(* IEC 61131-3 sources: JingjiangArm/moonboxpro_arm_8.4/Application/Application/任务列表/CommTask/COMM_DIAMONDS/和金刚UDP通讯/功能接口, 6 files *)

(* ---- KS_CheckAll_StZone_UnSynchronized.st ---- *)
(*@CES
Name=KS_CheckAll_StZone_UnSynchronized
Type=FunctionBlock
TypeGuid=6f9dac99-8de1-4efc-8465-68ac443b7d08
Guid=07bfdfe8-2771-43fc-9a3c-80039394908a
HasDeclaration=True
HasImplementation=True
*)
{DECLARATION}
FUNCTION KS_CheckAll_StZone_UnSynchronized : INT(*0表示都同步了/>0表示未同步的数量/<0表示错误*)
VAR_INPUT
	i_pstStDataZone: POINTER TO StDataZone;(*读写区域*)
END_VAR
VAR
	uiN: UINT;
	iResult: INT;
END_VAR

{IMPLEMENTATION}
iResult:= 0;
IF i_pstStDataZone<>0 THEN
	FOR uiN:=1 TO i_pstStDataZone^.uiNodeNum BY 1 DO
		IF i_pstStDataZone^.astStDataNode[uiN].bySynchronized<>SINT_TO_BYTE(-1) THEN
			iResult:= iResult+1;(*未同步的数量+1*)
		END_IF
	END_FOR
ELSE
	iResult:= -1;
END_IF
KS_CheckAll_StZone_UnSynchronized:= iResult;

(* ---- KS_GenTxData_.st ---- *)
(*@CES
Name=KS_GenTxData_
Type=FunctionBlock
TypeGuid=6f9dac99-8de1-4efc-8465-68ac443b7d08
Guid=4f0cddb0-57bc-4748-9ef3-99d0df4ac11d
HasDeclaration=True
HasImplementation=True
*)
{DECLARATION}
FUNCTION KS_GenTxData_ : INT(*0无错误/-1参数非法/-100未支持的功能字/-200写多个寄存器范围无效*)
VAR_INPUT
	i_dwTxBuf: DWORD;
	i_pstStDataNode: POINTER TO StDataNode;
	i_dwBaseAdr: DWORD;
	i_uiInvocation: UINT;
	i_byFunctionId: BYTE;(*功能id/目前仅处理03和16*)
	i_piTxPayloadLen: POINTER TO INT;(*用于接收返回的实际tx数据数量/单位字节*)
	i_xOnlyWrite: BOOL;(*只写区域-16384*)
END_VAR
VAR
	iResult: INT := 0;
	uiTmp: UINT;
	pstStADU_tmp: POINTER TO StADU;
	pbyByteCount_tmp: POINTER TO BYTE;
	paiRegisters_tmp: POINTER TO ARRAY [1..MAX_PDU_REGISTERS] OF INT;
END_VAR
VAR CONSTANT
	MAX_PDU_REGISTERS: INT := 123;(*0X1~0X7B(最大)*)
	MB_FUNC_READ_MULTI_REGS: BYTE := 3;(*读多个寄存器*)
	MB_FUNC_WRITE_MULTI_REGS: BYTE := 16;(*写多个寄存器*)
END_VAR
{IMPLEMENTATION}
iResult:= 0;
IF i_dwTxBuf<>0 AND
	i_pstStDataNode<>0 AND
	i_piTxPayloadLen<>0 THEN

	(*主要的输入参数合法*)
	pstStADU_tmp:= i_dwTxBuf;

	(*mbap*)
	pstStADU_tmp^.stStMBAP.uiInvocation:= bswap_16(i_uiInvocation);
	pstStADU_tmp^.stStMBAP.uiProtocol:= 0;
	pstStADU_tmp^.stStMBAP.uiLength:= 0;(*这个长度根据i_byFunctionId的类别最后再重新统计比较合适*)
	pstStADU_tmp^.stStMBAP.byUnit:= 1;(*按slaveID=1/2025.8.4.192327*)

	(*pdu*)
	pstStADU_tmp^.stStPDU_Header.byFunction:= i_byFunctionId;
	IF i_byFunctionId=MB_FUNC_READ_MULTI_REGS THEN(*读多个寄存器*)
		(*功能字/单字节/不需要字序处理*)
		pstStADU_tmp^.stStPDU_Header.byFunction:= i_byFunctionId;

		(*地址和寄存器数量/16bit/都需要做字序处理*)
		pstStADU_tmp^.stStPDU_Header.uiAddress:= bswap_16(i_pstStDataNode^.uiAddress);
		pstStADU_tmp^.stStPDU_Header.uiQuantity:= bswap_16(i_pstStDataNode^.uiQuantity);

		(*更新mbap中的uiLength/16bit/需要处理字序*)
		uiTmp:= SIZEOF(pstStADU_tmp^.stStMBAP.byUnit) + SIZEOF(pstStADU_tmp^.stStPDU_Header);
		pstStADU_tmp^.stStMBAP.uiLength:= bswap_16(uiTmp);

		(*实际数据量*)
		i_piTxPayloadLen^:= DWORD_TO_INT(SIZEOF(pstStADU_tmp^));

	ELSIF i_byFunctionId=MB_FUNC_WRITE_MULTI_REGS THEN(*写多个寄存器*)
		(*功能字/单字节/不需要字序处理*)
		pstStADU_tmp^.stStPDU_Header.byFunction:= i_byFunctionId;

		(*地址和寄存器数量/16bit/都需要做字序处理*)
		IF i_pstStDataNode^.uiQuantity>=1 AND i_pstStDataNode^.uiQuantity<=MAX_PDU_REGISTERS THEN
			(*增加1级判断/保证寄存器在合法范围*)

			pstStADU_tmp^.stStPDU_Header.uiAddress:= bswap_16(i_pstStDataNode^.uiAddress);
			pstStADU_tmp^.stStPDU_Header.uiQuantity:= bswap_16(i_pstStDataNode^.uiQuantity);

			(*填充字节数量/单字节不用做字序处理*)
			pbyByteCount_tmp:= i_dwTxBuf + SIZEOF(pstStADU_tmp^);
			pbyByteCount_tmp^:= UINT_TO_BYTE(i_pstStDataNode^.uiQuantity*2);

			(*将寄存器数据搬到要发送的区域/这里没有做大小端数据处理*)
			paiRegisters_tmp:= i_dwTxBuf + SIZEOF(pstStADU_tmp^) + SIZEOF(pbyByteCount_tmp^);
			IF i_xOnlyWrite THEN
				SysMemCpy(
					paiRegisters_tmp,
					i_dwBaseAdr+(i_pstStDataNode^.uiAddress-PARAM_ZONE_C2S)*2,
					i_pstStDataNode^.uiQuantity*2);
			ELSE
				SysMemCpy(
					paiRegisters_tmp,
					i_dwBaseAdr+(i_pstStDataNode^.uiAddress-PARAM_ZONE_ALTERNATE_OFST)*2,
					i_pstStDataNode^.uiQuantity*2);
			END_IF

			(*更新mbap中的uiLength/16bit/需要处理字序*)
			uiTmp:= SIZEOF(pstStADU_tmp^.stStMBAP.byUnit) + SIZEOF(pstStADU_tmp^.stStPDU_Header) + SIZEOF(pbyByteCount_tmp^) + i_pstStDataNode^.uiQuantity*2;
			pstStADU_tmp^.stStMBAP.uiLength:= bswap_16(uiTmp);

			(*实际数据量*)
			i_piTxPayloadLen^:= DWORD_TO_INT(SIZEOF(pstStADU_tmp^) + SIZEOF(pbyByteCount_tmp^) + i_pstStDataNode^.uiQuantity*2);
		ELSE
			iResult:= -200;
		END_IF
	ELSE
		iResult:= -100;(*未支持的功能字*)
	END_IF
ELSE
	iResult:= -1;
END_IF
KS_GenTxData_:= iResult;

(* ---- KS_InitStProofList.st ---- *)
(*@CES
Name=KS_InitStProofList
Type=FunctionBlock
TypeGuid=6f9dac99-8de1-4efc-8465-68ac443b7d08
Guid=42c94ff1-daf9-4f57-bbca-92a4069f4f99
HasDeclaration=True
HasImplementation=True
*)
{DECLARATION}
FUNCTION KS_InitStProofList : INT
VAR_INPUT
	i_pstStProofList: POINTER TO StProofList;
END_VAR
VAR
	iN: int;
	iResult: INT;
END_VAR

{IMPLEMENTATION}
iResult:= 0;
IF i_pstStProofList<>0 THEN
	(*清除证据链列表*)
	FOR iN:=1 TO MAX_MB_FIFO_ITEMS BY 1 DO
		i_pstStProofList^.astStProofItem[iN].iWaitRespCycles:= 0;
		i_pstStProofList^.astStProofItem[iN].stStADU.stStMBAP.uiInvocation:= 0;
		i_pstStProofList^.astStProofItem[iN].stStADU.stStMBAP.uiProtocol:= 0;
		i_pstStProofList^.astStProofItem[iN].stStADU.stStMBAP.uiLength:= 0;
		i_pstStProofList^.astStProofItem[iN].stStADU.stStMBAP.byUnit:= 0;
		i_pstStProofList^.astStProofItem[iN].stStADU.stStPDU_Header.byFunction:= 0;
		i_pstStProofList^.astStProofItem[iN].stStADU.stStPDU_Header.uiAddress:= 0;
		i_pstStProofList^.astStProofItem[iN].stStADU.stStPDU_Header.uiQuantity:= 0;
	END_FOR
ELSE
	iResult:= -1;
END_IF
KS_InitStProofList:= iResult;

(* ---- KS_InitStZone.st ---- *)
(*@CES
Name=KS_InitStZone
Type=FunctionBlock
TypeGuid=6f9dac99-8de1-4efc-8465-68ac443b7d08
Guid=6a7c2e7c-7aa2-44cc-96e1-c1f696e3ee98
HasDeclaration=True
HasImplementation=True
*)
{DECLARATION}
FUNCTION KS_InitStZone : INT(*0表示无错误/bit0置位表示读写区域错误/bit1置位表示只写区域错误*)
VAR_INPUT
	i_pstStParam_Diamonds_WrRd: POINTER TO StParam_Diamonds_WrRd;(*读写区域数据地址*)
	i_pstStDataZone_RW: POINTER TO StDataZone;(*读写区域*)
	i_pstStParam_Diamonds_Wr: POINTER TO StParam_Diamonds_Wr;(*只写区域数据地址*)
	i_pstStDataZone_W: POINTER TO StDataZone;(*只写区域*)
END_VAR
VAR
	iN: INT;
	iResult: INT;
	dwDlen: DWORD;
	dwBlocklen: DWORD;
	uiAddress: UINT;
END_VAR

{IMPLEMENTATION}
iResult:= 0;

(*读写区域*)
IF i_pstStParam_Diamonds_WrRd<>0 AND i_pstStDataZone_RW<>0 THEN
	i_pstStDataZone_RW^.uiNodeNum:= 0;
	dwDlen:= SIZEOF(i_pstStParam_Diamonds_WrRd^);
	dwBlocklen:= REGS_PER_DATA_NODE*2;
	uiAddress:= PARAM_ZONE_ALTERNATE_OFST;
	WHILE dwDlen>=dwBlocklen DO
		i_pstStDataZone_RW^.uiNodeNum:= i_pstStDataZone_RW^.uiNodeNum+1;
		i_pstStDataZone_RW^.astStDataNode[i_pstStDataZone_RW^.uiNodeNum].uiAddress:= uiAddress;
		i_pstStDataZone_RW^.astStDataNode[i_pstStDataZone_RW^.uiNodeNum].uiQuantity:= DWORD_TO_UINT(dwBlocklen/2);
		i_pstStDataZone_RW^.astStDataNode[i_pstStDataZone_RW^.uiNodeNum].bySynchronized:= 0;

		(*2025.8.5.094540/han.dp/+*)
		i_pstStDataZone_RW^.astStDataNode[i_pstStDataZone_RW^.uiNodeNum].xRd_ing:= FALSE;
		i_pstStDataZone_RW^.astStDataNode[i_pstStDataZone_RW^.uiNodeNum].xWr_ing:= FALSE;

		uiAddress:= uiAddress + i_pstStDataZone_RW^.astStDataNode[i_pstStDataZone_RW^.uiNodeNum].uiQuantity;
		dwDlen:= dwDlen-dwBlocklen;
	END_WHILE
	IF dwDlen>0 THEN
		i_pstStDataZone_RW^.uiNodeNum:= i_pstStDataZone_RW^.uiNodeNum+1;
		i_pstStDataZone_RW^.astStDataNode[i_pstStDataZone_RW^.uiNodeNum].uiAddress:= uiAddress;
		i_pstStDataZone_RW^.astStDataNode[i_pstStDataZone_RW^.uiNodeNum].uiQuantity:= DWORD_TO_UINT(dwDlen/2);
		i_pstStDataZone_RW^.astStDataNode[i_pstStDataZone_RW^.uiNodeNum].bySynchronized:= 0;

		(*2025.8.5.094540/han.dp/+*)
		i_pstStDataZone_RW^.astStDataNode[i_pstStDataZone_RW^.uiNodeNum].xRd_ing:= FALSE;
		i_pstStDataZone_RW^.astStDataNode[i_pstStDataZone_RW^.uiNodeNum].xWr_ing:= FALSE;
	END_IF
ELSE
	iResult:= iResult+1;
END_IF

(*只写区域*)
IF i_pstStParam_Diamonds_Wr<>0 AND i_pstStDataZone_W<>0 THEN
	i_pstStDataZone_W^.uiNodeNum:= 0;

	dwDlen:= SIZEOF(i_pstStParam_Diamonds_Wr^);
	dwBlocklen:= REGS_PER_DATA_NODE*2;
	uiAddress:= PARAM_ZONE_C2S;
	WHILE dwDlen>=dwBlocklen DO
		i_pstStDataZone_W^.uiNodeNum:= i_pstStDataZone_W^.uiNodeNum+1;
		i_pstStDataZone_W^.astStDataNode[i_pstStDataZone_W^.uiNodeNum].uiAddress:= uiAddress;
		i_pstStDataZone_W^.astStDataNode[i_pstStDataZone_W^.uiNodeNum].uiQuantity:= DWORD_TO_UINT(dwBlocklen/2);
		i_pstStDataZone_W^.astStDataNode[i_pstStDataZone_W^.uiNodeNum].bySynchronized:= 0;

		(*2025.8.5.094540/han.dp/+*)
		i_pstStDataZone_W^.astStDataNode[i_pstStDataZone_W^.uiNodeNum].xRd_ing:= FALSE;
		i_pstStDataZone_W^.astStDataNode[i_pstStDataZone_W^.uiNodeNum].xWr_ing:= FALSE;

		uiAddress:= uiAddress + i_pstStDataZone_W^.astStDataNode[i_pstStDataZone_W^.uiNodeNum].uiQuantity;
		dwDlen:= dwDlen-dwBlocklen;
	END_WHILE
	IF dwDlen>0 THEN
		i_pstStDataZone_W^.uiNodeNum:= i_pstStDataZone_W^.uiNodeNum+1;
		i_pstStDataZone_W^.astStDataNode[i_pstStDataZone_W^.uiNodeNum].uiAddress:= uiAddress;
		i_pstStDataZone_W^.astStDataNode[i_pstStDataZone_W^.uiNodeNum].uiQuantity:= DWORD_TO_UINT(dwDlen/2);
		i_pstStDataZone_W^.astStDataNode[i_pstStDataZone_W^.uiNodeNum].bySynchronized:= 0;

		(*2025.8.5.094540/han.dp/+*)
		i_pstStDataZone_W^.astStDataNode[i_pstStDataZone_W^.uiNodeNum].xRd_ing:= FALSE;
		i_pstStDataZone_W^.astStDataNode[i_pstStDataZone_W^.uiNodeNum].xWr_ing:= FALSE;
	END_IF

	iResult:= iResult+2;
END_IF

KS_InitStZone:= iResult;

(* ---- KS_PushDataToFifo.st ---- *)
(*@CES
Name=KS_PushDataToFifo
Type=FunctionBlock
TypeGuid=6f9dac99-8de1-4efc-8465-68ac443b7d08
Guid=b493b00e-9b49-48fd-b986-2a847e7b8547
HasDeclaration=True
HasImplementation=True
*)
{DECLARATION}
FUNCTION KS_PushDataToFifo : INT(*-1表示错误/>0表示写入的值数量/限制单次写入量1020有效内容*)
VAR_INPUT
	i_xRTdata: BOOL;(*TRUE表示‘RT'类型/FALSE表示'FI'类型*)
	i_pbyMem: POINTER TO BYTE;
	i_iBytesNum: INT;
	i_pstStUdpOnlySendFifo: POINTER TO StUdpOnlySendFifo;
END_VAR
VAR
	iResult: INT:= 0;
	byIdx_w: BYTE;
END_VAR

{IMPLEMENTATION}
iResult:= 0;
IF i_pbyMem<>0 AND
	i_iBytesNum>0 AND
	i_pstStUdpOnlySendFifo<>0 THEN
	(*参数合法*)

	byIdx_w:= i_pstStUdpOnlySendFifo^.byW;
	IF i_xRTdata THEN
		i_pstStUdpOnlySendFifo^.astStUdpOnlySend[byIdx_w].uiPkgTyp:= 16#5254;
	ELSE
		i_pstStUdpOnlySendFifo^.astStUdpOnlySend[byIdx_w].uiPkgTyp:= 16#4649;
	END_IF

	iResult:= MIN(SIZEOF(i_pstStUdpOnlySendFifo^.astStUdpOnlySend[byIdx_w].abyMem), i_iBytesNum);
	i_pstStUdpOnlySendFifo^.astStUdpOnlySend[byIdx_w].uiDlen:= INT_TO_UINT(iResult);

	SysMemCpy(
		ADR(i_pstStUdpOnlySendFifo^.astStUdpOnlySend[byIdx_w].abyMem),
		i_pbyMem,
		i_pstStUdpOnlySendFifo^.astStUdpOnlySend[byIdx_w].uiDlen);
	byIdx_w:= byIdx_w+1;
	i_pstStUdpOnlySendFifo^.byW:= byIdx_w;

ELSE
	iResult:= -1;
END_IF
KS_PushDataToFifo:= iResult;

(* ---- KS_Reset_StZone_SynchronizedFlag.st ---- *)
(*@CES
Name=KS_Reset_StZone_SynchronizedFlag
Type=FunctionBlock
TypeGuid=6f9dac99-8de1-4efc-8465-68ac443b7d08
Guid=96d189e0-34ee-41cd-a72d-4921ed0a61dc
HasDeclaration=True
HasImplementation=True
*)
{DECLARATION}
FUNCTION KS_Reset_StZone_SynchronizedFlag : INT
VAR_INPUT
	i_pstStDataZone: POINTER TO StDataZone;(*读写区域*)
END_VAR
VAR
	uiN: UINT;
	iResult: INT;
END_VAR

{IMPLEMENTATION}
iResult:= 0;
IF i_pstStDataZone<>0 THEN
	FOR uiN:=1 TO i_pstStDataZone^.uiNodeNum BY 1 DO
		i_pstStDataZone^.astStDataNode[uiN].bySynchronized:= 0;

		(*2025.8.5.094713/han.dp/如果写就置xWr_ing有效/如果读就置xRd_ing有效*)
		i_pstStDataZone^.astStDataNode[uiN].xRd_ing:= FALSE;
		i_pstStDataZone^.astStDataNode[uiN].xWr_ing:= FALSE;
	END_FOR
ELSE
	iResult:= -1;
END_IF
KS_Reset_StZone_SynchronizedFlag:= iResult;
